KUKA KRL program: MAIN_1.src

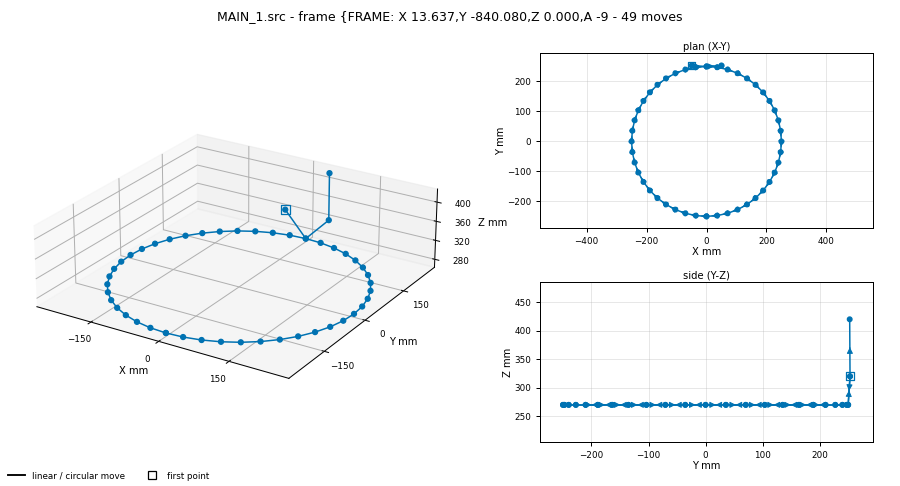
[picture p0: tool path of MAIN_1.src in frame {FRAME: X 13.637,Y -840.080,Z 0.000,A -9, 49 of 74 moves have a stored position in this frame; points joined in program order, loops and branches not executed]
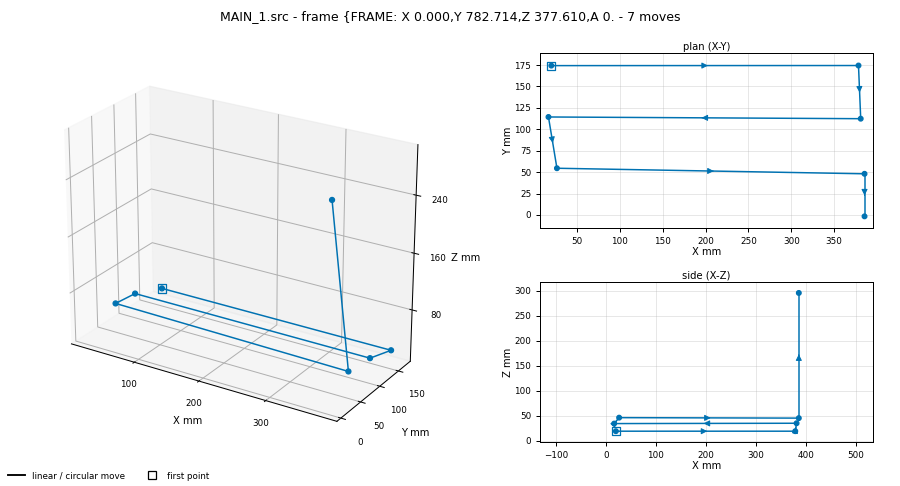
[picture p1: tool path of MAIN_1.src in frame {FRAME: X 0.000,Y 782.714,Z 377.610,A 0., 7 of 74 moves have a stored position in this frame; points joined in program order, loops and branches not executed]
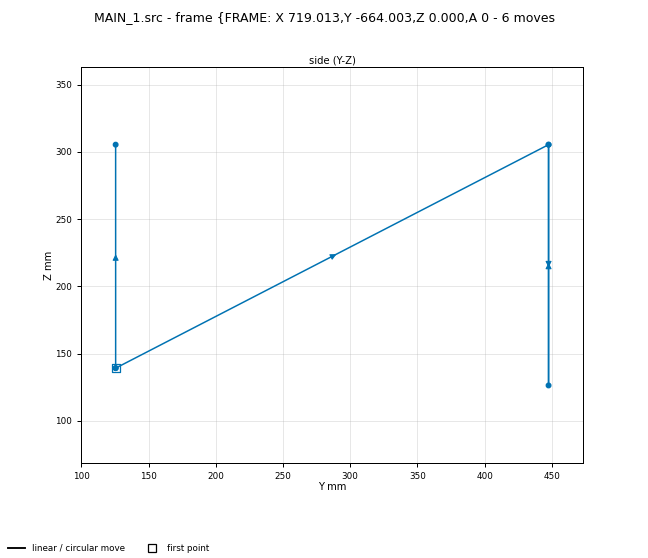
[picture p2: tool path of MAIN_1.src in frame {FRAME: X 719.013,Y -664.003,Z 0.000,A 0, 6 of 74 moves have a stored position in this frame; points joined in program order, loops and branches not executed]
&ACCESS RVP
&REL 1
&PARAM TEMPLATE = C:\KRC\Roboter\Template\vorgabe
&PARAM EDITMASK = *
DEF MAIN_1 ( )

; External program calls:
EXT REMOTE_PROG_CALL()
EXT PICK_PART_111()
EXT PLACE_PART_112()
EXT EVENT_PROG_START()
EXT EVENT_PATH_APPRO()
EXT EVENT_PATH_START()
EXT EVENT_PATH_FINIS()
EXT EVENT_PATH_RETRA()
EXT EVENT_PROG_FINIS()
EXT PROG_1___with_a_()

EXT BAS (BAS_COMMAND :IN,REAL :IN )


; GLOBAL INTERRUPT DECL 3 WHEN $STOPMESS==TRUE DO IR_STOPM ( )
; INTERRUPT ON 3

;FOLD Initialise and set default speed
BAS (#INITMOV,0)
BAS (#VEL_PTP,100)
BAS (#ACC_PTP,20)
$VEL.CP=0.2
BAS (#TOOL,0)
BAS (#BASE,0)
;ENDFOLD

;;FOLD STARTPOS
;$BWDSTART = FALSE
;PDAT_ACT = PDEFAULT
;BAS(#PTP_DAT)
;FDAT_ACT = {TOOL_NO 0,BASE_NO 0,IPO_FRAME #BASE}
;BAS(#FRAMES)
;;ENDFOLD

$ADVANCE = 5

;FOLD ---- Quickly skip BCO ----
; PTP $AXIS_ACT
;ENDFOLD

;FOLD ---- GO HOME ----
; PTP {A1 0.000, A2 -90.000, A3 90.000, A4 0.000, A5 0.000, A6 0.000, E1 0, E2 0, E3 0, E4 0, E5 0, E6 0}
;ENDFOLD


; Program generated by RoboDK v5.6.9 for RoboDK Industrial on 26/02/2024 09:58:20
; Using nominal kinematics.
PTP {A1 -0.00000,A2 0.00000,A3 0.00000,A4 0.00000,A5 0.00000,A6 -0.00000,E1 0.00000}
PTP {A1 0.00000,A2 3.21124,A3 -15.42370,A4 0.00000,A5 12.21250,A6 -0.00000,E1 0.00000}
LIN {X 1015.000,Y 0.000,Z 1272.000,A 0.000,B 90.000,C 0.000,E1 0.00000, S 'B110', T 'B0010100'}
$OUT[5]=TRUE
$OUT[5]=TRUE
$OUT[5]=0.5
$OUT[5]=true
$ANOUT[5]=TRUE
$ANOUT[5]=TRUE
$ANOUT[5]=0.5
$ANOUT[5]=true
var=val
var=val
WAIT FOR ($IN[5]==TRUE)
WAIT FOR ($IN[5]==TRUE)
WAIT FOR ($IN[5]==0.5)
WAIT FOR ($IN[5]==true)
START_TIMER:
$TIMER_STOP[1]=TRUE
$TIMER_FLAG[1]=FALSE
$TIMER[1]=0.100
$TIMER_STOP[1]=FALSE
WAIT FOR ($IN[5]==TRUE OR $TIMER_FLAG[1])
$TIMER_STOP[1]=TRUE
IF $TIMER_FLAG[1]== TRUE THEN
    HALT ; Timed out!
    GOTO START_TIMER
ENDIF
WAIT FOR (var==val)
START_TIMER:
$TIMER_STOP[1]=TRUE
$TIMER_FLAG[1]=FALSE
$TIMER[1]=0.100
$TIMER_STOP[1]=FALSE
WAIT FOR (var==val OR $TIMER_FLAG[1])
$TIMER_STOP[1]=TRUE
IF $TIMER_FLAG[1]== TRUE THEN
    HALT ; Timed out!
    GOTO START_TIMER
ENDIF
Wait for StrClear($LOOP_MSG[])
$LOOP_CONT = TRUE
$LOOP_MSG[] = "Message"
REMOTE_PROG_CALL()
CODE_INSERT_172
; Insert Comment
; ---- Setting reference (Base) ----
$BASE = {FRAME: X 719.013,Y -664.003,Z 0.000,A 0.000,B 0.000,C 0.000}
; --------------------------
; ---- Setting tool (TCP) ----
; TOOL_DATA[1] = {FRAME: X 129.073,Y 0.000,Z 85.477,A 0.000,B 22.849,C 0.000}
$TOOL = {FRAME: X 129.073,Y 0.000,Z 85.477,A 0.000,B 22.849,C 0.000}
; $TOOL = TOOL_DATA[1]
; --------------------------
$ACC.ORI1 = 800.00000
$ACC.ORI2 = 800.00000
$VEL.ORI1 = 500.00000
$VEL.ORI2 = 500.00000
$APO.CPTP = 10
$APO.CDIS = 10.000
PTP {A1 -29.33220,A2 46.67700,A3 -0.02452,A4 26.54560,A5 25.39570,A6 -51.63400,E1 0.00000} C_PTP
$ACC.CP = 0.20000
$VEL.CP = 0.10000
LIN {X 187.786,Y 125.499,Z 139.112,A -179.997,B 0.180,C 179.996,E1 0.00000, S 'B010', T 'B0100101'}
$OUT[5]=TRUE
PICK_PART_111()
$APO.CPTP = 10
$APO.CDIS = 10.000
$ACC.CP = 0.60000
$VEL.CP = 0.30000
; Linear movement using joint targets is not supported. Change the target type to cartesian or use a joint movement.
LIN {X 187.272,Y 447.522,Z 305.347,A 179.999,B 0.185,C -179.998,E1 0.00000, S 'B010', T 'B0100001'} C_DIS
$ACC.CP = 0.20000
$VEL.CP = 0.10000
; MoveSearch command not implemented
LIN {X 187.851,Y 447.517,Z 126.235,A 179.999,B 0.185,C -179.998,E1 0.00000, S 'B010', T 'B0100001'}
$OUT[5]=FALSE
PLACE_PART_112()
$APO.CPTP = 10
$APO.CDIS = 10.000
LIN {X 187.272,Y 447.522,Z 305.347,A 179.999,B 0.185,C -179.998,E1 0.00000, S 'B010', T 'B0100001'} C_DIS
; ---- Setting reference (Base) ----
$BASE = {FRAME: X 577.670,Y 392.250,Z 0.000,A 38.960,B 0.000,C 0.000}
; --------------------------
$APO.CPTP = 25
$APO.CDIS = 25.000
$ACC.ORI1 = 800.00000
$ACC.ORI2 = 800.00000
$VEL.ORI1 = 500.00000
$VEL.ORI2 = 500.00000
$ACC.CP = 0.20000
$VEL.CP = 0.10000
PTP {A1 52.18600,A2 45.67580,A3 6.92000,A4 66.73420,A5 19.93230,A6 -92.73000,E1 0.00000} C_PTP
CIRC {X 430.047,Y 43.774,Z 231.503,A -134.549,B 11.181,C 178.913 S 'B010', T 'B100100'},{X 109.688,Y -153.222,Z 161.073,A -134.549,B 11.181,C 178.913,E1 0.00000 S 'B010', T 'B0100000'} C_DIS
; Circular movement using joint targets is not supported. Change the target type to cartesian or use a joint movement.
$ACC.CP = 0.20000
$VEL.CP = 0.10000
LIN {X 312.208,Y 292.214,Z 255.156,A -134.549,B 11.181,C 178.913,E1 0.00000, S 'B010', T 'B0100000'}
PTP {A1 -0.00000,A2 0.00000,A3 0.00000,A4 0.00000,A5 0.00000,A6 -0.00000,E1 0.00000}
; ---- Setting reference (Base) ----
$BASE = {FRAME: X 0.000,Y 782.714,Z 377.610,A 0.000,B 0.000,C 0.000}
; --------------------------
PTP {A1 88.67600,A2 29.60160,A3 -6.42883,A4 -1.98422,A5 49.47920,A6 4.54769,E1 0.00000}
LIN {X 19.898,Y 174.307,Z 19.008,A -94.928,B -5.426,C -179.533,E1 0.00000, S 'B010', T 'B0001000'}
LIN {X 378.402,Y 174.416,Z 18.997,A -94.928,B -5.426,C -179.533,E1 0.00000, S 'B010', T 'B0100100'}
LIN {X 380.996,Y 112.363,Z 34.882,A -95.294,B -18.136,C -178.348,E1 0.00000, S 'B010', T 'B0101000'}
LIN {X 16.551,Y 114.359,Z 34.226,A -95.294,B -18.136,C -178.348,E1 0.00000, S 'B010', T 'B0001000'}
LIN {X 26.434,Y 54.524,Z 46.072,A -95.461,B 4.348,C 179.585,E1 0.00000, S 'B010', T 'B0001000'}
LIN {X 385.448,Y 48.050,Z 45.137,A -95.590,B 11.181,C 178.913,E1 0.00000, S 'B010', T 'B0100000'}
LIN {X 385.448,Y -1.625,Z 295.251,A -95.590,B 11.181,C 178.913,E1 0.00000, S 'B010', T 'B0100000'}
PTP {A1 -0.00000,A2 0.00000,A3 0.00000,A4 0.00000,A5 0.00000,A6 -0.00000,E1 0.00000}
EVENT_PROG_START()
$APO.CPTP = 1
$APO.CDIS = 1.000
$VEL.CP = 1.00000
; ---- Setting reference (Base) ----
$BASE = {FRAME: X 13.637,Y -840.080,Z 0.000,A -90.000,B 0.000,C 0.000}
; --------------------------
; Show Tool 1
PTP {A1 -68.09030,A2 24.20190,A3 26.78550,A4 38.21340,A5 36.20170,A6 -98.79640,E1 0.00000} C_PTP
EVENT_PATH_APPRO()
LIN {X -49.895,Y 253.259,Z 319.999,A -90.000,B 0.353,C -179.975,E1 0.00000, S 'B010', T 'B0100001'} C_DIS
LIN {X 0.000,Y 250.000,Z 270.000,A -90.000,B 0.353,C -179.975,E1 0.00000, S 'B010', T 'B0100001'} C_DIS
EVENT_PATH_START()
$VEL.CP = 0.05000
LIN {X 35.579,Y 247.455,Z 270.000,A -90.000,B 0.345,C -179.925,E1 0.00000, S 'B010', T 'B0100001'} C_DIS
LIN {X 70.433,Y 239.873,Z 270.000,A -89.999,B 0.331,C -179.876,E1 0.00000, S 'B010', T 'B0100001'} C_DIS
LIN {X 103.854,Y 227.408,Z 270.000,A -89.999,B 0.310,C -179.831,E1 0.00000, S 'B010', T 'B0100001'} C_DIS
LIN {X 135.160,Y 210.313,Z 270.000,A -89.999,B 0.283,C -179.788,E1 0.00000, S 'B010', T 'B0100001'} C_DIS
LIN {X 163.715,Y 188.937,Z 270.000,A -89.999,B 0.250,C -179.750,E1 0.00000, S 'B010', T 'B0100001'} C_DIS
LIN {X 188.937,Y 163.715,Z 270.000,A -89.999,B 0.212,C -179.717,E1 0.00000, S 'B010', T 'B0100001'} C_DIS
LIN {X 210.313,Y 135.160,Z 270.000,A -89.999,B 0.170,C -179.689,E1 0.00000, S 'B010', T 'B0100001'} C_DIS
LIN {X 227.408,Y 103.854,Z 270.000,A -89.999,B 0.124,C -179.668,E1 0.00000, S 'B010', T 'B0100001'} C_DIS
LIN {X 239.873,Y 70.433,Z 270.000,A -90.000,B 0.075,C -179.654,E1 0.00000, S 'B010', T 'B0100001'} C_DIS
LIN {X 247.455,Y 35.579,Z 270.000,A -90.000,B 0.025,C -179.647,E1 0.00000, S 'B010', T 'B0100001'} C_DIS
LIN {X 250.000,Y 0.000,Z 270.000,A -90.000,B -0.025,C -179.647,E1 0.00000, S 'B010', T 'B0100001'} C_DIS
LIN {X 247.455,Y -35.579,Z 270.000,A -90.000,B -0.075,C -179.654,E1 0.00000, S 'B010', T 'B0100001'} C_DIS
LIN {X 239.873,Y -70.433,Z 270.000,A -90.001,B -0.124,C -179.668,E1 0.00000, S 'B010', T 'B0100001'} C_DIS
LIN {X 227.408,Y -103.854,Z 270.000,A -90.001,B -0.170,C -179.689,E1 0.00000, S 'B010', T 'B0100001'} C_DIS
LIN {X 210.313,Y -135.160,Z 270.000,A -90.001,B -0.212,C -179.717,E1 0.00000, S 'B010', T 'B0100001'} C_DIS
LIN {X 188.937,Y -163.715,Z 270.000,A -90.001,B -0.250,C -179.750,E1 0.00000, S 'B010', T 'B0100001'} C_DIS
LIN {X 163.715,Y -188.937,Z 270.000,A -90.001,B -0.283,C -179.788,E1 0.00000, S 'B010', T 'B0100001'} C_DIS
LIN {X 135.160,Y -210.313,Z 270.000,A -90.001,B -0.311,C -179.830,E1 0.00000, S 'B010', T 'B0100001'} C_DIS
LIN {X 103.854,Y -227.408,Z 270.000,A -90.001,B -0.332,C -179.876,E1 0.00000, S 'B010', T 'B0100001'} C_DIS
LIN {X 70.433,Y -239.873,Z 270.000,A -90.000,B -0.346,C -179.925,E1 0.00000, S 'B010', T 'B0100001'} C_DIS
LIN {X 35.579,Y -247.455,Z 270.000,A -90.000,B -0.353,C -179.975,E1 0.00000, S 'B010', T 'B0100001'} C_DIS
LIN {X 0.000,Y -250.000,Z 270.000,A -90.000,B -0.353,C -179.975,E1 0.00000, S 'B010', T 'B0100001'} C_DIS
LIN {X 0.000,Y -250.000,Z 270.000,A -90.000,B -0.353,C 179.975,E1 0.00000, S 'B010', T 'B0100001'} C_DIS
LIN {X -35.579,Y -247.455,Z 270.000,A -90.000,B -0.346,C 179.925,E1 0.00000, S 'B010', T 'B0100001'} C_DIS
LIN {X -70.433,Y -239.873,Z 270.000,A -89.999,B -0.331,C 179.876,E1 0.00000, S 'B010', T 'B0100001'} C_DIS
LIN {X -103.854,Y -227.408,Z 270.000,A -89.999,B -0.310,C 179.831,E1 0.00000, S 'B010', T 'B0100001'} C_DIS
LIN {X -135.160,Y -210.313,Z 270.000,A -89.999,B -0.283,C 179.788,E1 0.00000, S 'B010', T 'B0100001'} C_DIS
LIN {X -163.715,Y -188.937,Z 270.000,A -89.999,B -0.250,C 179.750,E1 0.00000, S 'B010', T 'B0100001'} C_DIS
LIN {X -188.937,Y -163.715,Z 270.000,A -89.999,B -0.212,C 179.717,E1 0.00000, S 'B010', T 'B0100001'} C_DIS
LIN {X -210.313,Y -135.160,Z 270.000,A -89.999,B -0.169,C 179.690,E1 0.00000, S 'B010', T 'B0100001'} C_DIS
LIN {X -227.408,Y -103.854,Z 270.000,A -89.999,B -0.123,C 179.669,E1 0.00000, S 'B010', T 'B0100001'} C_DIS
LIN {X -239.873,Y -70.433,Z 270.000,A -90.000,B -0.075,C 179.654,E1 0.00000, S 'B010', T 'B0100001'} C_DIS
LIN {X -247.455,Y -35.579,Z 270.000,A -90.000,B -0.025,C 179.647,E1 0.00000, S 'B010', T 'B0100001'} C_DIS
LIN {X -250.000,Y 0.000,Z 270.000,A -90.000,B 0.025,C 179.647,E1 0.00000, S 'B010', T 'B0100001'} C_DIS
LIN {X -247.455,Y 35.579,Z 270.000,A -90.000,B 0.075,C 179.655,E1 0.00000, S 'B010', T 'B0100001'} C_DIS
LIN {X -239.873,Y 70.433,Z 270.000,A -90.001,B 0.123,C 179.669,E1 0.00000, S 'B010', T 'B0100001'} C_DIS
LIN {X -227.408,Y 103.854,Z 270.000,A -90.001,B 0.170,C 179.689,E1 0.00000, S 'B010', T 'B0100001'} C_DIS
LIN {X -210.313,Y 135.160,Z 270.000,A -90.001,B 0.212,C 179.717,E1 0.00000, S 'B010', T 'B0100001'} C_DIS
LIN {X -188.937,Y 163.715,Z 270.000,A -90.001,B 0.250,C 179.750,E1 0.00000, S 'B010', T 'B0100001'} C_DIS
LIN {X -163.715,Y 188.937,Z 270.000,A -90.001,B 0.283,C 179.788,E1 0.00000, S 'B010', T 'B0100001'} C_DIS
LIN {X -135.160,Y 210.313,Z 270.000,A -90.001,B 0.310,C 179.831,E1 0.00000, S 'B010', T 'B0100001'} C_DIS
LIN {X -103.854,Y 227.408,Z 270.000,A -90.001,B 0.332,C 179.876,E1 0.00000, S 'B010', T 'B0100001'} C_DIS
LIN {X -70.433,Y 239.873,Z 270.000,A -90.000,B 0.346,C 179.925,E1 0.00000, S 'B010', T 'B0100001'} C_DIS
LIN {X -35.579,Y 247.455,Z 270.000,A -90.000,B 0.353,C 179.975,E1 0.00000, S 'B010', T 'B0100001'} C_DIS
LIN {X 0.000,Y 250.000,Z 270.000,A -90.000,B 0.353,C 179.975,E1 0.00000, S 'B010', T 'B0100001'} C_DIS
$VEL.CP = 1.00000
EVENT_PATH_FINIS()
LIN {X 49.895,Y 253.258,Z 319.999,A -90.000,B 0.353,C 179.975,E1 0.00000, S 'B010', T 'B0100001'} C_DIS
LIN {X 49.939,Y 252.642,Z 419.997,A -90.000,B 0.353,C 179.975,E1 0.00000, S 'B010', T 'B0100001'} C_DIS
EVENT_PATH_RETRA()
EVENT_PROG_FINIS()
; ---- Setting reference (Base) ----
$BASE = {FRAME: X 719.013,Y -664.003,Z 0.000,A 0.000,B 0.000,C 0.000}
; --------------------------
PTP {A1 -29.33220,A2 46.67700,A3 -0.02452,A4 26.54560,A5 25.39570,A6 -51.63400,E1 0.00000} C_PTP
WAIT SEC 1.250
LIN {X 187.786,Y 125.499,Z 139.112,A -179.997,B 0.180,C 179.996,E1 0.00000, S 'B010', T 'B0100101'} C_DIS
WAIT FOR ($IN[1]==TRUE)
LIN {X 187.264,Y 125.487,Z 305.356,A 180.000,B 0.184,C -180.000,E1 0.00000, S 'B010', T 'B0100101'} C_DIS
PROG_1___with_a_()
END
